// TIA Portal V20 export
Screen "200PRBCompleteDisplay"  1276x673
  ScreenItem "sequenceControlFaceplate_Lite_1" at 392,556 size 641x64  Type=HmiFaceplateContainer
  ScreenItem "Title_ScreenOverview_X390_Y2" at 390,2 size 500x30  Type=HmiTextBox
  ScreenItem "Button_Back_1" at 2,2 size 90x60  Type=HmiButton
  ScreenItem "Line_Header_X0_Y64" at 0,64 size 1276x0  Type=HmiLine
  ScreenItem "Tec-Unit_LegendᆉY2" at 1183,2 size 90x60  Type=HmiButton
  ScreenItem "permanentareaborderrectangle" at 0,0 size 0x0  Type=HmiRectangle
  ScreenItem "Button_Back" at 2,4 size 90x60  Type=HmiButton
  ScreenItem "Title_ScreenOverview_X390_Y2_1" at 380,5 size 510x57  Type=HmiTextBox
  ScreenItem "面板容器_1" at 10,267 size 163x70  Type=HmiFaceplateContainer
  ScreenItem "面板容器_3" at 196,334 size 163x70  Type=HmiFaceplateContainer
  ScreenItem "面板容器_4" at 10,335 size 163x70  Type=HmiFaceplateContainer
  ScreenItem "面板容器_5" at 619,334 size 163x70  Type=HmiFaceplateContainer
  ScreenItem "面板容器_6" at 431,267 size 163x70  Type=HmiFaceplateContainer
  ScreenItem "面板容器_7" at 431,335 size 163x70  Type=HmiFaceplateContainer
  ScreenItem "面板容器_8" at 848,335 size 163x70  Type=HmiFaceplateContainer
  ScreenItem "面板容器_9" at 1048,267 size 163x70  Type=HmiFaceplateContainer
  ScreenItem "面板容器_10" at 848,267 size 163x70  Type=HmiFaceplateContainer
  ScreenItem "面板容器_11" at 10,605 size 163x70  Type=HmiFaceplateContainer
  ScreenItem "面板容器_12" at 431,605 size 163x70  Type=HmiFaceplateContainer
  ScreenItem "面板容器_13" at 848,605 size 163x70  Type=HmiFaceplateContainer
  ScreenItem "面板容器_2" at 1090,4 size 88x58  Type=HmiFaceplateContainer
  ScreenItem "OPMode1_Blocked" at 1164,6 size 14x14  Type=HmiGraphicView
  ScreenItem "OPMode4_Foreground_Blocked_1" at 1090,4 size 88x58  Type=HmiGraphicView
  ScreenItem "Button_Back_2" at 1180,606 size 90x60  Type=HmiButton
  ScreenItem "面板容器_14" at 196,267 size 163x70  Type=HmiFaceplateContainer
  ScreenItem "面板容器_15" at 619,267 size 163x70  Type=HmiFaceplateContainer
